Fanuc KAREL source: KT00930.KL

PROGRAM KT00930
%NOLOCKGROUP
VAR
  R1: REAL
  R2: REAL
  OUT: INTEGER
BEGIN
  R1 = 2.0
  R2 = 3.0
  R1 = 2.0
  R2 = 3.0
  OUT = ORD(R1, 1)
END KT00930
